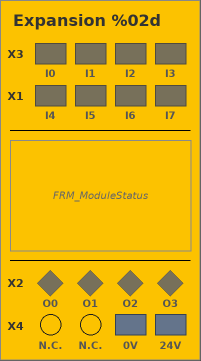
VISUALIZATION FRM_Module8DI4DO  // 201x361
VAR_IN_OUT
   stModuleData: ST_PNOZModuleData;
END_VAR
VAR_INPUT
   nIndex: USINT;  
END_VAR
    Rectangle (0,0 201x361)
    Line (10,130) (190,130)
    Line (10,260) (190,260)
    Label (0,44 31x21), "X3"
    Label (0,86 31x21), "X1"
    Label (0,273 31x21), "X2"
    Label (0,316 31x21), "X4"
    Frame (10,140 181x111)
        shows FRM_ModuleStatus(bPower := stModuleData.stLEDState.bPower, bRun := stModuleData.stLEDState.bRun, bDiag := stModuleData.stLEDState.bDiag, bFault := stModuleData.stLEDState.bFault, bInputFault := stModuleData.stLEDState.bInputFault, bOutputFault := stModuleData.stLEDState.bOutputFault, sName := stModuleData.sName, nID := stModuleData.nID, nSerialNumber := stModuleData.nSerialNumber, anRevision := stModuleData.anDeviceVersion)
    Textfield (10,0 181x41), "Expansion %02d", text variable: nIndex
    Label (30,68 41x11), "I0"
    Label (70,68 41x11), "I1"
    Label (110,68 41x11), "I2"
    Label (150,68 41x11), "I3"
    Label (30,110 41x11), "I4"
    Label (70,110 41x11), "I5"
    Label (110,110 41x11), "I6"
    Label (150,110 41x11), "I7"
    Label (30,298 41x11), "O0"
    Label (70,298 41x11), "O1"
    Label (110,298 41x11), "O2"
    Label (150,298 41x11), "O3"
    Label (30,340 41x11), "N.C."
    Label (70,340 41x11), "N.C."
    Label (110,340 41x11), "0V"
    Label (150,340 41x11), "24V"
    Ellipse (40,314 21x21)
    Ellipse (80,314 21x21)
    Rectangle (115,314 31x21)
    Rectangle (155,314 31x21)
    Rectangle (35,43 31x21), colour toggle: stModuleData.anInput[1].b0
    Rectangle (75,43 31x21), colour toggle: stModuleData.anInput[1].b1
    Rectangle (115,43 31x21), colour toggle: stModuleData.anInput[1].b2
    Rectangle (155,43 31x21), colour toggle: stModuleData.anInput[1].b3
    Rectangle (35,85 31x21), colour toggle: stModuleData.anInput[1].b4
    Rectangle (75,85 31x21), colour toggle: stModuleData.anInput[1].b5
    Rectangle (115,85 31x21), colour toggle: stModuleData.anInput[1].b6
    Rectangle (155,85 31x21), colour toggle: stModuleData.anInput[1].b7
    Polygon (37,283) (50,270) (63,283) (50,296) (50,296), colour toggle: stModuleData.anOutput[1].b0
    Polygon (77,283) (90,270) (103,283) (90,296) (90,296), colour toggle: stModuleData.anOutput[1].b1
    Polygon (117,283) (130,270) (143,283) (130,296) (130,296), colour toggle: stModuleData.anOutput[1].b2
    Polygon (157,283) (170,270) (183,283) (170,296) (170,296), colour toggle: stModuleData.anOutput[1].b3
END_VISUALIZATION

(* stored: Version 1.1.0.1
   Visu FRM_Module8DI4DO: Id {576eab5a-5fc3-05e7-2c47-1fa1883ecb05} *)
